Fanuc KAREL source: KO00108.KL

PROGRAM KO00108
%NOLOCKGROUP
VAR
  A: REAL
  B: REAL
  OUT: REAL
BEGIN
  A = 1
  B = 2
  OUT = ATAN2(A, B)
END KO00108
